Staubli VAL3: stop.pgx

program stop()
// Stop motion and carriage; preserve vacuum command.
begin
  // ============================================================
  // PARADA SIN SOLTAR AUTOMATICAMENTE UNA PIEZA
  // ============================================================
  resetMotion()
  trolleyOn = false
  barrierClosed = true
  // TODO FISICO: confirmar que barrierClosed=true realmente cierra bOut5.
  // vacuumOn se conserva para no soltar una pieza al ordenar STOP.
  cycleOK = false
  cycleStep = -1
  putln("Stopped: inspect station before restarting")
end
